{attribute 'Tc2GvlVarNames'}
VAR_GLOBAL
	stgGr01Alarm			:ST_AlarmRef;
END_VAR

(* stored: Version 1.1.0.1, ProductVersion 3.1.4024.15
   GVL GVL_Gr01Alarm: Id {e859b2f7-e709-435d-8a2f-da2f55ee14da} *)
